SUBAPPLICATION Klappen_Sitzventile (* Subapplication Type *)
  (* Standard: 61499-2 *)
  (* Version 1.0, 2023-02-11, franz *)
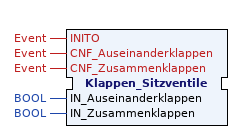
  EVENT_INPUT
    INITO;
    CNF_Auseinanderklappen;
    CNF_Zusammenklappen;
  END_EVENT
  VAR_INPUT
    IN_Auseinanderklappen : BOOL;
    IN_Zusammenklappen : BOOL;
  END_VAR
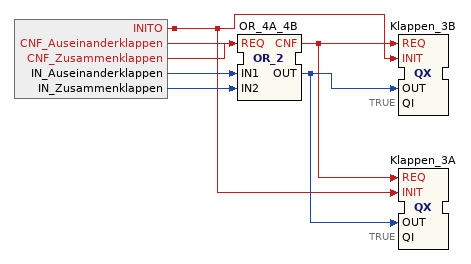
  FBS
    OR_4A_4B : OR_2; {SET_ATTRIBUTE(PinComment, IN1:Auseinanderklappen)} {SET_ATTRIBUTE(PinComment, IN2:Zusammenklappen)}
    Klappen_3B : QX(QI := TRUE);
    Klappen_3A : QX(QI := TRUE);
  END_FBS
  EVENT_CONNECTIONS
    OR_4A_4B.CNF TO Klappen_3B.REQ;
    OR_4A_4B.CNF TO Klappen_3A.REQ;
    CNF_Auseinanderklappen TO OR_4A_4B.REQ;
    CNF_Zusammenklappen TO OR_4A_4B.REQ;
    INITO TO Klappen_3B.INIT;
    INITO TO Klappen_3A.INIT;
  END_CONNECTIONS
  DATA_CONNECTIONS
    OR_4A_4B.OUT TO Klappen_3B.OUT;
    OR_4A_4B.OUT TO Klappen_3A.OUT;
    IN_Auseinanderklappen TO OR_4A_4B.IN1;
    IN_Zusammenklappen TO OR_4A_4B.IN2;
  END_CONNECTIONS
END_SUBAPPLICATION
